Staubli VAL3: utText.dtx

public string sFontFamily
public string sFontStyle
public num nFontSize
